# EPICS substitutions: db/Beckhoff_7XXX/ecmcEP7041-3102.substitutions
file "ecmcEL7037-chX.template"
{
  pattern {CH_ID}
          {01   }
}

file "ecmcEL5101-chX.template"
{
  pattern {CH_ID}
          {01   }
}
